FUNCTION_BLOCK SortingOwnership (* Sorting-only architecture following Distribution and tutorial modules 1-4 *)
  (* Standard: 61499-2 *)
  (* Version 2.0, 2026-11-09, sorting2n, sorting2n *)
  PACKAGE Main;
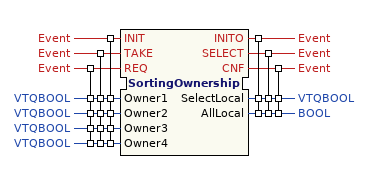
  EVENT_INPUT
    INIT WITH Owner1, Owner2, Owner3, Owner4;
    TAKE WITH Owner1, Owner2, Owner3, Owner4;
    REQ WITH Owner1, Owner2, Owner3, Owner4;
  END_EVENT
  EVENT_OUTPUT
    INITO WITH SelectLocal, AllLocal;
    SELECT WITH SelectLocal, AllLocal;
    CNF WITH SelectLocal, AllLocal;
  END_EVENT
  VAR_INPUT
    Owner1 : VTQBOOL;
    Owner2 : VTQBOOL;
    Owner3 : VTQBOOL;
    Owner4 : VTQBOOL;
  END_VAR
  VAR_OUTPUT
    SelectLocal : VTQBOOL;
    AllLocal : BOOL;
  END_VAR
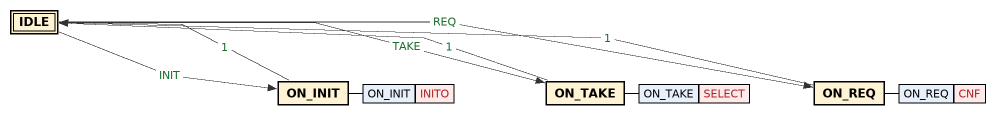
  EC_STATES
    IDLE;
    ON_INIT : ON_INIT -> INITO;
    ON_TAKE : ON_TAKE -> SELECT;
    ON_REQ : ON_REQ -> CNF;
  END_STATES
  EC_TRANSITIONS
    IDLE TO ON_INIT := INIT;
    ON_INIT TO IDLE := 1;
    IDLE TO ON_TAKE := TAKE;
    ON_TAKE TO IDLE := 1;
    IDLE TO ON_REQ := REQ;
    ON_REQ TO IDLE := 1;
  END_TRANSITIONS
  ALGORITHM ON_INIT IN ST:
SelectLocal.value := FALSE; SelectLocal.quality := 0; AllLocal := FALSE;
  END_ALGORITHM
  ALGORITHM ON_TAKE IN ST:
SelectLocal.value := TRUE; SelectLocal.quality := 0;
  END_ALGORITHM
  ALGORITHM ON_REQ IN ST:
AllLocal := Owner1.value AND Owner2.value AND Owner3.value AND Owner4.value;
  END_ALGORITHM
END_FUNCTION_BLOCK
